(* IEC 61131-3 sources: MappView1/ECTempSim/ECTempSim, 3 files *)

(* ---- ECTempSim.typ ---- *)
(********************************************************************
 * COPYRIGHT -- Bernecker + Rainer
 ********************************************************************
 * Library: TempLib
 * File: TempLib.typ
 * Author: gierlingerj
 * Created: May 15, 2013
 ********************************************************************
 * Data types of library TempLib
 ********************************************************************)

TYPE
	SimModInternalType : 	STRUCT
		Tt_cool : MTBasicsTimeDelay;
		Tt_heat : MTBasicsTimeDelay;
		PT2 : MTBasicsPT2;
		k_h : REAL := 1.0;
		k_c : REAL := 1.0;
		EnableOld : BOOL;
		RoomTemp : REAL;
	END_STRUCT;
END_TYPE

(* ---- ECTempSim.fun ---- *)
(********************************************************************
 * COPYRIGHT -- Bernecker + Rainer
 ********************************************************************
 * Library: TempLib
 * File: TempLib.fun
 * Author: gierlingerj
 * Created: May 15, 2013
 ********************************************************************
 * Functions and function blocks of library TempLib
 ********************************************************************)

FUNCTION_BLOCK ECTempSimModel (*simulation of an extruder temperature zone*) (*$GROUP=User*)
	VAR_INPUT
		Enable : BOOL; (*Enables the function block*)
		InHeat : REAL; (*Heating control action. Permitted values: 0.0..100.0 [%].*)
		InCool : REAL; (*Cooling control action. Permitted values: 0.0..100.0 [%].*)
	END_VAR
	VAR_OUTPUT
		Active : BOOL; (*Function block is active.*)
		Error : BOOL; (*Indicates an error.*)
		StatusID : UDINT; (*Status information.*)
		UpdateDone : BOOL; (*Update is done.*)
		OutTemp : REAL; (*Output temperature (output variable). Units: °C.*)
	END_VAR
	VAR
		Internal : SimModInternalType;
	END_VAR
END_FUNCTION_BLOCK

(* ---- ECTempSim.var ---- *)
(********************************************************************
 * COPYRIGHT -- Bernecker + Rainer
 ********************************************************************
 * Library: TempLib
 * File: TempLib.var
 * Author: gierlingerj
 * Created: May 15, 2013
 ********************************************************************
 * Constants of library TempLib
 ********************************************************************)
VAR CONSTANT
	ERR_TEMPLIB_GAIN_INVALID : DINT := 45000;
	ERR_TEMPLIB_TUNING_RANGE_INVALID : DINT := 50000;
END_VAR
